KUKA KRL program: Main_Program.src

&ACCESS RVP
&REL 1
&PARAM TEMPLATE = C:\KRC\Roboter\Template\vorgabe
&PARAM EDITMASK = *
DEF Main_Program ( )

; External program calls:
EXT Home_Motoman()
EXT Home_KUKA()
EXT Drilling()
EXT Chamfer()
EXT Paint()
EXT onDrilling_Start()
EXT onDrilling_Appro()
EXT onDrilling_PathS()
EXT onDrilling_Activ()
EXT onDrilling_Retra()
EXT onDrilling_Finis()
EXT onChamfer_Start()
EXT onChamfer_Approa()
EXT onChamfer_PathSt()
EXT onChamfer_Retrac()
EXT onChamfer_Finish()
EXT onPaint_Start()
EXT SetRPM()
EXT onPaint_Approach()
EXT onPaint_PathStar()
EXT onPaint_Retract()
EXT onPaint_Finish()

EXT BAS (BAS_COMMAND :IN,REAL :IN )


; GLOBAL INTERRUPT DECL 3 WHEN $STOPMESS==TRUE DO IR_STOPM ( )
; INTERRUPT ON 3

;FOLD Initialise and set default speed
BAS (#INITMOV,0)
BAS (#VEL_PTP,100)
BAS (#ACC_PTP,20)
$VEL.CP=0.2
BAS (#TOOL,0)
BAS (#BASE,0)
;ENDFOLD

;;FOLD STARTPOS
;$BWDSTART = FALSE
;PDAT_ACT = PDEFAULT
;BAS(#PTP_DAT)
;FDAT_ACT = {TOOL_NO 0,BASE_NO 0,IPO_FRAME #BASE}
;BAS(#FRAMES)
;;ENDFOLD

$ADVANCE = 5

;FOLD ---- Quickly skip BCO ----
; PTP $AXIS_ACT
;ENDFOLD

;FOLD ---- GO HOME ----
; PTP {A1 0.000, A2 -90.000, A3 90.000, A4 0.000, A5 0.000, A6 0.000, E1 0, E2 0, E3 0, E4 0, E5 0, E6 0}
;ENDFOLD


; Program generated by VerticalBot Studio for KUKA KR 90 R3100 extra on 25/10/2026 12:00:00
; Using nominal kinematics.
; ---- Setting reference (Base) ----
; BASE_DATA[1] = {FRAME: X 1545.530,Y 599.115,Z 1469.820,A 93.801,B 0.000,C 0.000}
$BASE = {FRAME: X 1545.530,Y 599.115,Z 1469.820,A 93.801,B 0.000,C 0.000}
; $BASE = BASE_DATA[1]
; --------------------------
; ---- Setting tool (TCP) ----
$TOOL = {FRAME: X 260.000,Y 0.000,Z 292.000,A 0.000,B 90.000,C 0.000}
; --------------------------
WAIT SEC 5.000
Home_Motoman()
Home_KUKA()
Drilling()
Chamfer()
Paint()
Home_Motoman()
Home_KUKA()
WAIT SEC 5.000
END
